Staubli VAL3: addLog.pgx

public program addLog(string x_sLog (dimensions=1), num x_nType (dimensions=1))
begin
  call Log:addlog(x_sLog,x_nType)
end
